FUNCTION_BLOCK FT_TEST
VAR_INPUT
  CLK : BOOL;
END_VAR
VAR
  f : F_TRIG;
END_VAR
BEGIN
  f(CLK := CLK);
  //#ASSERT NOT f.Q : Pbad
END_FUNCTION_BLOCK
